// TIA Portal V20 export
Screen "RobotCollision"  1276x673
  ScreenItem "Title_ScreenOverview_X390_Y2" at 438,5 size 510x57  Type=HmiTextBox
  ScreenItem "Line_Header_X0_Y64" at 0,64 size 1274x1  Type=HmiLine
  ScreenItem "矩形_6" at 6,69 size 1262x597  Type=HmiRectangle
  ScreenItem "permanentareaborderrectangle" at 0,0 size 0x0  Type=HmiRectangle
  ScreenItem "Button_Back" at 2,2 size 90x60  Type=HmiButton
  ScreenItem "Graphic view_1" at 225,-96 size 744x865  Type=HmiGraphicView
  ScreenItem "Graphic view_4" at 596,199 size 147x35  Type=HmiGraphicView
  ScreenItem "Graphic view_2" at 595,149 size 153x35  Type=HmiGraphicView
  ScreenItem "Text_1" at 637,107 size 88x35  Type=HmiText
  ScreenItem "Text_2" at 884,183 size 88x35  Type=HmiText
  ScreenItem "Text_3" at 884,532 size 88x35  Type=HmiText
  ScreenItem "Text_4" at 334,532 size 88x35  Type=HmiText
  ScreenItem "Text_5" at 334,184 size 88x35  Type=HmiText
  ScreenItem "Text_6" at 637,246 size 88x35  Type=HmiText
  ScreenItem "Graphic view_3" at 595,510 size 153x35  Type=HmiGraphicView
  ScreenItem "Graphic view_5" at 596,560 size 147x35  Type=HmiGraphicView
  ScreenItem "Text_7" at 637,468 size 88x35  Type=HmiText
  ScreenItem "Text_8" at 637,607 size 88x35  Type=HmiText
  ScreenItem "Rectangle_2" at 8,5 size 164x111  Type=HmiRectangle
  ScreenItem "Text_13" at 0,0 size 174x35  Type=HmiText
  ScreenItem "Text_14" at 31,26 size 123x35  Type=HmiText
  ScreenItem "Text_15" at 44,54 size 88x35  Type=HmiText
  ScreenItem "Text_16" at 37,82 size 136x35  Type=HmiText
  ScreenItem "矩形_7" at 21,89 size 17x17  Type=HmiRectangle
  ScreenItem "矩形_5" at 21,62 size 17x17  Type=HmiRectangle
  ScreenItem "矩形_4" at 21,35 size 17x17  Type=HmiRectangle
  ScreenItem "Rectangle_7" at 8,5 size 161x111  Type=HmiRectangle
  ScreenItem "Text_33" at 0,0 size 171x35  Type=HmiText
  ScreenItem "Text_34" at 32,26 size 121x35  Type=HmiText
  ScreenItem "Text_35" at 45,54 size 87x35  Type=HmiText
  ScreenItem "Text_36" at 38,82 size 134x35  Type=HmiText
  ScreenItem "矩形_20" at 18,35 size 17x17  Type=HmiRectangle
  ScreenItem "矩形_21" at 18,62 size 17x17  Type=HmiRectangle
  ScreenItem "矩形_22" at 18,89 size 17x17  Type=HmiRectangle
  ScreenItem "Rectangle_1" at 8,5 size 164x111  Type=HmiRectangle
  ScreenItem "Text_9" at 0,0 size 174x35  Type=HmiText
  ScreenItem "Text_10" at 31,26 size 123x35  Type=HmiText
  ScreenItem "Text_11" at 44,54 size 88x35  Type=HmiText
  ScreenItem "Text_12" at 37,82 size 136x35  Type=HmiText
  ScreenItem "矩形_10" at 20,89 size 17x17  Type=HmiRectangle
  ScreenItem "矩形_9" at 20,62 size 17x17  Type=HmiRectangle
  ScreenItem "矩形_8" at 20,35 size 17x17  Type=HmiRectangle
  ScreenItem "Rectangle_6" at 8,5 size 164x111  Type=HmiRectangle
  ScreenItem "Text_29" at 0,0 size 174x35  Type=HmiText
  ScreenItem "Text_30" at 31,26 size 123x35  Type=HmiText
  ScreenItem "Text_31" at 44,54 size 88x35  Type=HmiText
  ScreenItem "Text_32" at 37,82 size 136x35  Type=HmiText
  ScreenItem "矩形_1" at 20,35 size 17x17  Type=HmiRectangle
  ScreenItem "矩形_2" at 20,62 size 17x17  Type=HmiRectangle
  ScreenItem "矩形_3" at 20,89 size 17x17  Type=HmiRectangle
